Fanuc KAREL source: NC0069.KL

-- PROVISIONAL review KL for V940-1; original PC SHA256 0760343ee36e4ab3a756b061e1f3dfcda60b747224ea0bda51b71d62ef0fae9c
-- Incomplete behavior may be omitted. Consult companion uncertainty JSON. Do not deploy.
PROGRAM NC0069
%NOLOCKGROUP
-- UNRESOLVED_LOCAL_POOL 16 cells at code offset 3; source declarations unknown
-- DIRECT_LOCAL_WORD_ACCESS alone does not prove INTEGER, REAL, or BOOLEAN
BEGIN
  -- V9_EXPOSED_INDEXED_TABLE_HINT layout=0001; 30 counted words exposed once; source arms/runtime held
  -- V9_FOOTER_20_HINT 15 numerical footer links; VM transfer unproved
  -- UNRESOLVED_PC offsets 0-8; opcodes 2B,2C,7B
  -- UNRESOLVED_PC offsets 13-20; opcodes 9D,23
  -- UNRESOLVED_PC offsets 25-54; opcodes 9D,23,9E,2E,22,7A
  -- UNRESOLVED_PC offsets 59-88; opcodes 9D,23,9E,2E,22,7A
  -- UNRESOLVED_PC offsets 93-122; opcodes 9D,23,9E,2E,22,7A
  -- UNRESOLVED_PC offsets 127-156; opcodes 9D,23,9E,2E,22,7A
  -- UNRESOLVED_PC offsets 161-190; opcodes 9D,23,9E,2E,22,7A
  -- UNRESOLVED_PC offsets 195-224; opcodes 9D,23,9E,2E,22,7A
  -- UNRESOLVED_PC offsets 229-258; opcodes 9D,23,9E,2E,22,7A
  -- UNRESOLVED_PC offsets 263-292; opcodes 9D,23,9E,2E,22,7A
  -- UNRESOLVED_PC offsets 297-326; opcodes 9D,23,9E,2E,22,7A
  -- UNRESOLVED_PC offsets 331-360; opcodes 9D,23,9E,2E,22,7A
  -- UNRESOLVED_PC offsets 365-394; opcodes 9D,23,9E,2E,22,7A
  -- UNRESOLVED_PC offsets 399-428; opcodes 9D,23,9E,2E,22,7A
  -- UNRESOLVED_PC offsets 433-462; opcodes 9D,23,9E,2E,22,7A
  -- UNRESOLVED_PC offsets 467-496; opcodes 9D,23,9E,2E,22,7A
  -- UNRESOLVED_PC offsets 501-530; opcodes 9D,23,9E,2E,22,7A
  -- UNRESOLVED_PC offsets 535-549; opcodes 21,9D,52,23
  -- UNRESOLVED_PC offsets 554-569; opcodes 20,2C,23
  -- UNRESOLVED_PC offsets 574-589; opcodes 20,2C,23
  -- UNRESOLVED_PC offsets 594-609; opcodes 20,2C,23
  -- UNRESOLVED_PC offsets 614-629; opcodes 20,2C,23
  -- UNRESOLVED_PC offsets 634-649; opcodes 20,2C,23
  -- UNRESOLVED_PC offsets 654-669; opcodes 20,2C,23
  -- UNRESOLVED_PC offsets 674-689; opcodes 20,2C,23
  -- UNRESOLVED_PC offsets 694-709; opcodes 20,2C,23
  -- UNRESOLVED_PC offsets 714-729; opcodes 20,2C,23
  -- UNRESOLVED_PC offsets 734-749; opcodes 20,2C,23
  -- UNRESOLVED_PC offsets 754-769; opcodes 20,2C,23
  -- UNRESOLVED_PC offsets 774-789; opcodes 20,2C,23
  -- UNRESOLVED_PC offsets 794-809; opcodes 20,2C,23
  -- UNRESOLVED_PC offsets 814-829; opcodes 20,2C,23
  -- UNRESOLVED_PC offsets 834-849; opcodes 20,2C,23
  -- UNRESOLVED_PC offsets 854-858; opcodes 7F
  -- UNRESOLVED_PC offsets 863-867; opcodes 27,AA
  -- UNRESOLVED_PC offsets 872-876; opcodes 7F
END NC0069
